(* IEC 61131-3 sources: plc-st-coding-agent/progress/evidence/f14_v6_public_pilot_20261112/jobs/codex_deepseek-v4pro (part 2) *)

(* ---- public-medium-04.raw_candidate_02.st ---- *)
FUNCTION_BLOCK FB
VAR_INPUT
    TemperatureSensorInput : REAL;
    SetTemperature : REAL;
END_VAR
VAR_OUTPUT
    CurrentTemperature : REAL;
    SetTempDisplay : REAL;
    HeaterStatus : BOOL;
    OverheatProtection : BOOL;
    HeaterOutput : BOOL;
END_VAR
VAR
    local_SensorFault : BOOL;
    local_HeatCommand : BOOL;
    local_OverheatActive : BOOL;
    HeaterContinuousTimer : TON;
    OverheatCooldownTimer : TON;
END_VAR

(*
ENGINEERING_CONTRACT
- Displays follow inputs each scan; REAL values are passed through without conversion (PUB002/PUB007).
- Normal heat: on when TemperatureSensorInput < SetTemperature; off when TemperatureSensorInput >= SetTemperature.
  Equality is unspecified by PUB003-PUB005 and is interpreted as off.
- Sensor fault: TemperatureSensorInput < 0.0 OR TemperatureSensorInput > 100.0 forces heat off.
  Values 0.0 and 100.0 remain valid (PUB008).
- Overheat: triggered only after continuous heating exceeds 5 s (strict > boundary implemented as
  T#5001MS). The trip starts a 3 s release timer; HeaterOutput remains off and OverheatProtection
  clears when the release timer reaches T#3S (PUB006).
- Same-scan priority: sensor fault / active overheat overrides normal demand; a continuous-heat
  timer trip overrides the computed heat command in that scan and starts the release timer.
- Units/boundaries: TIME uses T#5001MS for the heat trip and T#3S for release.
*)

(* CONTRACT_RULES [] *)

CurrentTemperature := TemperatureSensorInput;
SetTempDisplay := SetTemperature;

local_SensorFault := (TemperatureSensorInput < 0.0) OR (TemperatureSensorInput > 100.0);

IF local_SensorFault OR local_OverheatActive THEN
    local_HeatCommand := FALSE;
ELSIF TemperatureSensorInput < SetTemperature THEN
    local_HeatCommand := TRUE;
ELSE
    local_HeatCommand := FALSE;
END_IF;

HeaterContinuousTimer(IN := local_HeatCommand, PT := T#5001MS);
IF HeaterContinuousTimer.Q THEN
    local_OverheatActive := TRUE;
    local_HeatCommand := FALSE;
END_IF;

IF local_OverheatActive THEN
    OverheatCooldownTimer(IN := TRUE, PT := T#3S);
    IF OverheatCooldownTimer.Q THEN
        local_OverheatActive := FALSE;
    END_IF;
ELSE
    OverheatCooldownTimer(IN := FALSE, PT := T#3S);
END_IF;

HeaterOutput := local_HeatCommand AND NOT local_SensorFault AND NOT local_OverheatActive;
HeaterStatus := HeaterOutput;
OverheatProtection := local_OverheatActive;

END_FUNCTION_BLOCK

(* ---- public-medium-08.candidate_01.st ---- *)
FUNCTION_BLOCK FB_IPv4Parser
(* ENGINEERING_CONTRACT
   Output ipValue:
   - Activation: parsed and refreshed synchronously on every scan.
   - Hold: no latching; value is recomputed from ipText each scan.
   - Reset/deactivation: invalid input writes UDINT#0.
   - Same-scan priority: final overall validity wins over partial accumulation.
   - Units/bounds: UDINT 0..4294967295, segments 0..255.
   - Segment count/nonempty rules: PUB002, PUB004.
   - Byte order and assembly: PUB003, first byte at bits 24..31.
*)
(* CONTRACT_RULES [] *)
VAR_INPUT
    ipText : STRING(254);
END_VAR
VAR_OUTPUT
    ipValue : UDINT;
END_VAR
VAR
    tmp_i : INT;
    tmp_len : INT;
    tmp_ch : USINT;
    tmp_segCount : INT;
    tmp_segLen : INT;
    tmp_shift : INT;
    tmp_segValue : UDINT;
    tmp_result : UDINT;
    tmp_valid : BOOL;
END_VAR

ipValue := UDINT#0;
tmp_valid := TRUE;
tmp_segCount := 0;
tmp_segLen := 0;
tmp_segValue := UDINT#0;
tmp_result := UDINT#0;
tmp_len := LEN(ipText);

FOR tmp_i := 0 TO tmp_len - 1 DO
    tmp_ch := BYTE_TO_USINT(ipText[tmp_i]);

    IF tmp_ch = USINT#46 THEN
        IF tmp_segLen = 0 THEN
            tmp_valid := FALSE;
            EXIT;
        END_IF;

        tmp_segCount := tmp_segCount + 1;
        IF tmp_segCount > 4 THEN
            tmp_valid := FALSE;
            EXIT;
        END_IF;

        tmp_shift := (4 - tmp_segCount) * 8;
        tmp_result := tmp_result + SHL(tmp_segValue, tmp_shift);
        tmp_segLen := 0;
        tmp_segValue := UDINT#0;
    ELSIF (tmp_ch >= USINT#48) AND (tmp_ch <= USINT#57) THEN
        tmp_segLen := tmp_segLen + 1;
        tmp_segValue := tmp_segValue * UDINT#10
                        + (USINT_TO_UDINT(tmp_ch) - UDINT#48);

        IF tmp_segValue > UDINT#255 THEN
            tmp_valid := FALSE;
            EXIT;
        END_IF;
    ELSE
        tmp_valid := FALSE;
        EXIT;
    END_IF;
END_FOR;

IF tmp_valid AND (tmp_segLen > 0) THEN
    tmp_segCount := tmp_segCount + 1;

    IF tmp_segCount = 4 THEN
        tmp_result := tmp_result + tmp_segValue;
        ipValue := tmp_result;
    ELSE
        ipValue := UDINT#0;
    END_IF;
ELSE
    ipValue := UDINT#0;
END_IF;
END_FUNCTION_BLOCK

(* ---- public-medium-08.raw_candidate_01.st ---- *)
FUNCTION_BLOCK FB_IPv4Parser
(* ENGINEERING_CONTRACT
   Output ipValue:
   - Activation: parsed and refreshed synchronously on every scan.
   - Hold: no latching; value is recomputed from ipText each scan.
   - Reset/deactivation: invalid input writes UDINT#0.
   - Same-scan priority: final overall validity wins over partial accumulation.
   - Units/bounds: UDINT 0..4294967295, segments 0..255.
   - Segment count/nonempty rules: PUB002, PUB004.
   - Byte order and assembly: PUB003, first byte at bits 24..31.
*)
(* CONTRACT_RULES [] *)
VAR_INPUT
    ipText : STRING(254);
END_VAR
VAR_OUTPUT
    ipValue : UDINT;
END_VAR
VAR
    tmp_i : INT;
    tmp_len : INT;
    tmp_ch : USINT;
    tmp_segCount : INT;
    tmp_segLen : INT;
    tmp_shift : INT;
    tmp_segValue : UDINT;
    tmp_result : UDINT;
    tmp_valid : BOOL;
END_VAR

ipValue := UDINT#0;
tmp_valid := TRUE;
tmp_segCount := 0;
tmp_segLen := 0;
tmp_segValue := UDINT#0;
tmp_result := UDINT#0;
tmp_len := LEN(ipText);

FOR tmp_i := 0 TO tmp_len - 1 DO
    tmp_ch := BYTE_TO_USINT(ipText[tmp_i]);

    IF tmp_ch = USINT#46 THEN
        IF tmp_segLen = 0 THEN
            tmp_valid := FALSE;
            EXIT;
        END_IF;

        tmp_segCount := tmp_segCount + 1;
        IF tmp_segCount > 4 THEN
            tmp_valid := FALSE;
            EXIT;
        END_IF;

        tmp_shift := (4 - tmp_segCount) * 8;
        tmp_result := tmp_result + SHL(tmp_segValue, tmp_shift);
        tmp_segLen := 0;
        tmp_segValue := UDINT#0;
    ELSIF (tmp_ch >= USINT#48) AND (tmp_ch <= USINT#57) THEN
        tmp_segLen := tmp_segLen + 1;
        tmp_segValue := tmp_segValue * UDINT#10
                        + (USINT_TO_UDINT(tmp_ch) - UDINT#48);

        IF tmp_segValue > UDINT#255 THEN
            tmp_valid := FALSE;
            EXIT;
        END_IF;
    ELSE
        tmp_valid := FALSE;
        EXIT;
    END_IF;
END_FOR;

IF tmp_valid AND (tmp_segLen > 0) THEN
    tmp_segCount := tmp_segCount + 1;

    IF tmp_segCount = 4 THEN
        tmp_result := tmp_result + tmp_segValue;
        ipValue := tmp_result;
    ELSE
        ipValue := UDINT#0;
    END_IF;
ELSE
    ipValue := UDINT#0;
END_IF;
END_FUNCTION_BLOCK
